REGION Network 105: STATE Num:300 StChkTTPos
   RUNG wire#powerrail
      Contact( #s300_StChkTTPos )
      wire#w1
      I_Contact( #sStWtResetRel )
      I_Contact( #s300_StChkTTPos_T1 )
      I_Contact( #s300_StChkTTPos_T2 )
      I_Contact( #s300_StChkTTPos_T3 )
      wire#w2
      Coil( #s300_StChkTTPos )
   END_RUNG
   RUNG wire#powerrail
      Contact( #s20_StChkForPalletPresent_T4 )
   END_RUNG wire#w1
   RUNG wire#w2
      { S7_GenerateENO := "TRUE" } Move(in := 300, out1 => #StateNo)
   END_RUNG
   // the same network as SCL:
   #s300_StChkTTPos := (#s300_StChkTTPos OR #s20_StChkForPalletPresent_T4) AND NOT #sStWtResetRel AND NOT #s300_StChkTTPos_T1 AND NOT #s300_StChkTTPos_T2 AND NOT #s300_StChkTTPos_T3;
   IF #s300_StChkTTPos THEN #StateNo := 300; END_IF;
END_REGION

REGION Network 106: Actions for STATE Num:300 StChkTTPos
   RUNG wire#powerrail
      Contact( #s300_StChkTTPos )
      Coil( #qOutput1 )
   END_RUNG
   // the same network as SCL:
   #qOutput1 := #s300_StChkTTPos;
END_REGION

REGION Network 107: Transition for STATE Num:310 StWtRTRFrmTTUpAt0
   RUNG wire#powerrail
      Contact( #s310_StWtRTRFrmTTUpAt0 )
      I_Contact( #sStWtResetRel )
      Contact( #sSst )
      wire#w1
      Contact( #sTTUp_Timer_ON.Q )
      Coil( #s310_StWtRTRFrmTTUpAt0_T1 )
   END_RUNG
   RUNG wire#w1
      I_Contact( #s310_StWtRTRFrmTTUpAt0_T1 )
      Contact( #iOTS_Frm_Prev_TTUp )
      I_Contact( #sTTUp_Timer_ON.Q )
      Coil( #s310_StWtRTRFrmTTUpAt0_T2 )
   END_RUNG
   // the same network as SCL:
   #_w1 := #s310_StWtRTRFrmTTUpAt0 AND NOT #sStWtResetRel AND #sSst;
   #s310_StWtRTRFrmTTUpAt0_T1 := #_w1 AND #sTTUp_Timer_ON.Q;
   #s310_StWtRTRFrmTTUpAt0_T2 := #_w1 AND NOT #s310_StWtRTRFrmTTUpAt0_T1 AND #iOTS_Frm_Prev_TTUp AND NOT #sTTUp_Timer_ON.Q;
END_REGION

REGION Network 108: STATE Num:310 StWtRTRFrmTTUpAt0
   RUNG wire#powerrail
      Contact( #s310_StWtRTRFrmTTUpAt0 )
      wire#w1
      I_Contact( #sStWtResetRel )
      I_Contact( #s310_StWtRTRFrmTTUpAt0_T1 )
      I_Contact( #s310_StWtRTRFrmTTUpAt0_T2 )
      wire#w2
      Coil( #s310_StWtRTRFrmTTUpAt0 )
   END_RUNG
   RUNG wire#powerrail
      Contact( #s300_StChkTTPos_T1 )
   END_RUNG wire#w1
   RUNG wire#w2
      { S7_GenerateENO := "TRUE" } Move(in := 310, out1 => #StateNo)
   END_RUNG
   // the same network as SCL:
   #s310_StWtRTRFrmTTUpAt0 := (#s310_StWtRTRFrmTTUpAt0 OR #s300_StChkTTPos_T1) AND NOT #sStWtResetRel AND NOT #s310_StWtRTRFrmTTUpAt0_T1 AND NOT #s310_StWtRTRFrmTTUpAt0_T2;
   IF #s310_StWtRTRFrmTTUpAt0 THEN #StateNo := 310; END_IF;
END_REGION

REGION Network 109: Actions for STATE Num:310 StWtRTRFrmTTUpAt0
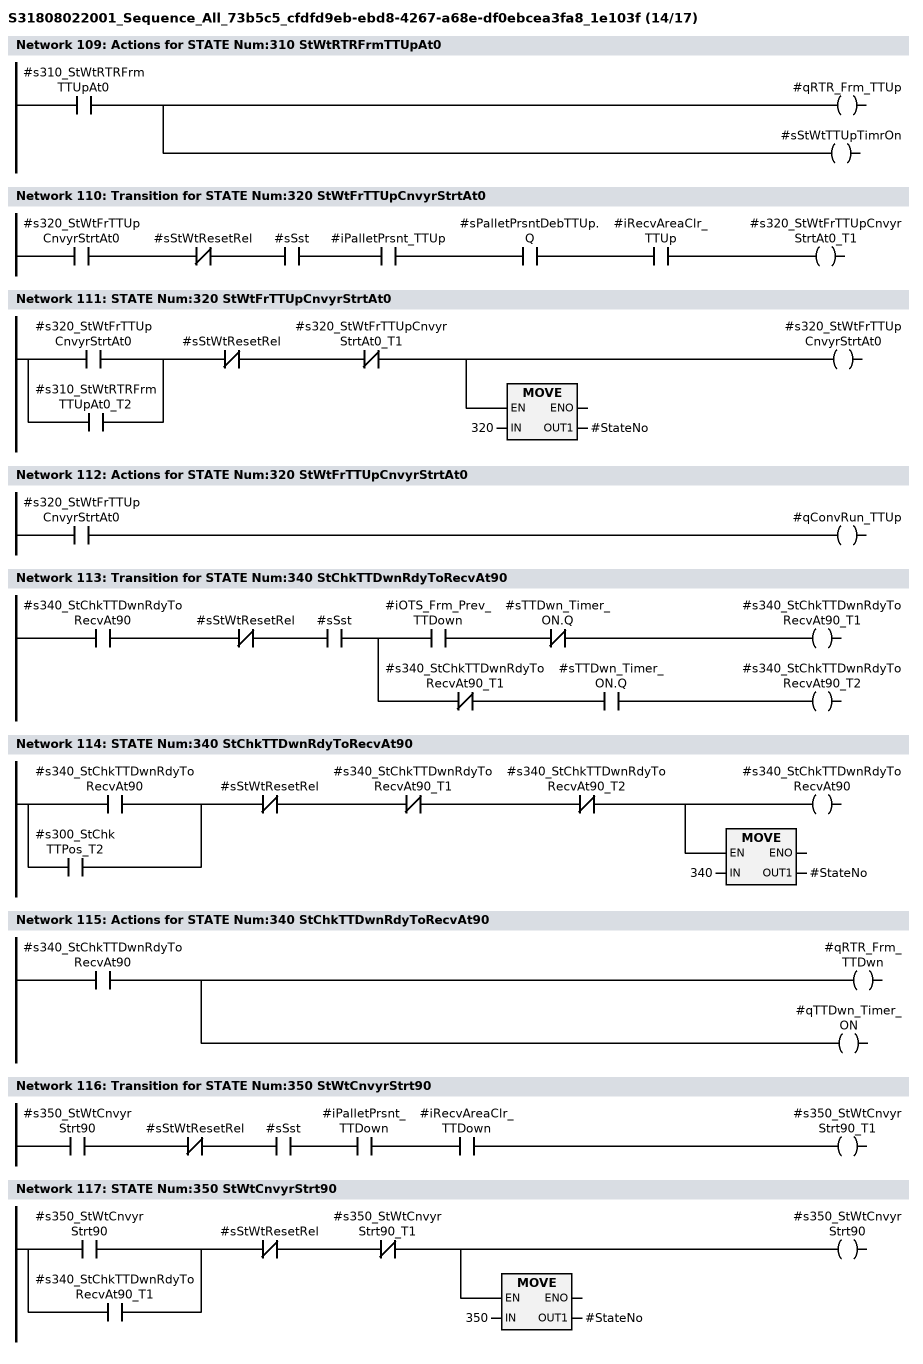
   RUNG wire#powerrail
      Contact( #s310_StWtRTRFrmTTUpAt0 )
      wire#w1
      Coil( #qRTR_Frm_TTUp )
   END_RUNG
   RUNG wire#w1
      Coil( #sStWtTTUpTimrOn )
   END_RUNG
   // the same network as SCL:
   #qRTR_Frm_TTUp := #s310_StWtRTRFrmTTUpAt0;
   #sStWtTTUpTimrOn := #s310_StWtRTRFrmTTUpAt0;
END_REGION

REGION Network 110: Transition for STATE Num:320 StWtFrTTUpCnvyrStrtAt0
   RUNG wire#powerrail
      Contact( #s320_StWtFrTTUpCnvyrStrtAt0 )
      I_Contact( #sStWtResetRel )
      Contact( #sSst )
      Contact( #iPalletPrsnt_TTUp )
      Contact( #sPalletPrsntDebTTUp.Q )
      Contact( #iRecvAreaClr_TTUp )
      Coil( #s320_StWtFrTTUpCnvyrStrtAt0_T1 )
   END_RUNG
   // the same network as SCL:
   #s320_StWtFrTTUpCnvyrStrtAt0_T1 := #s320_StWtFrTTUpCnvyrStrtAt0 AND NOT #sStWtResetRel AND #sSst AND #iPalletPrsnt_TTUp AND #sPalletPrsntDebTTUp.Q AND #iRecvAreaClr_TTUp;
END_REGION

REGION Network 111: STATE Num:320 StWtFrTTUpCnvyrStrtAt0
   RUNG wire#powerrail
      Contact( #s320_StWtFrTTUpCnvyrStrtAt0 )
      wire#w1
      I_Contact( #sStWtResetRel )
      I_Contact( #s320_StWtFrTTUpCnvyrStrtAt0_T1 )
      wire#w2
      Coil( #s320_StWtFrTTUpCnvyrStrtAt0 )
   END_RUNG
   RUNG wire#powerrail
      Contact( #s310_StWtRTRFrmTTUpAt0_T2 )
   END_RUNG wire#w1
   RUNG wire#w2
      { S7_GenerateENO := "TRUE" } Move(in := 320, out1 => #StateNo)
   END_RUNG
   // the same network as SCL:
   #s320_StWtFrTTUpCnvyrStrtAt0 := (#s320_StWtFrTTUpCnvyrStrtAt0 OR #s310_StWtRTRFrmTTUpAt0_T2) AND NOT #sStWtResetRel AND NOT #s320_StWtFrTTUpCnvyrStrtAt0_T1;
   IF #s320_StWtFrTTUpCnvyrStrtAt0 THEN #StateNo := 320; END_IF;
END_REGION

REGION Network 112: Actions for STATE Num:320 StWtFrTTUpCnvyrStrtAt0
   RUNG wire#powerrail
      Contact( #s320_StWtFrTTUpCnvyrStrtAt0 )
      Coil( #qConvRun_TTUp )
   END_RUNG
   // the same network as SCL:
   #qConvRun_TTUp := #s320_StWtFrTTUpCnvyrStrtAt0;
END_REGION

REGION Network 113: Transition for STATE Num:340 StChkTTDwnRdyToRecvAt90
   RUNG wire#powerrail
      Contact( #s340_StChkTTDwnRdyToRecvAt90 )
      I_Contact( #sStWtResetRel )
      Contact( #sSst )
      wire#w1
      Contact( #iOTS_Frm_Prev_TTDown )
      I_Contact( #sTTDwn_Timer_ON.Q )
      Coil( #s340_StChkTTDwnRdyToRecvAt90_T1 )
   END_RUNG
   RUNG wire#w1
      I_Contact( #s340_StChkTTDwnRdyToRecvAt90_T1 )
      Contact( #sTTDwn_Timer_ON.Q )
      Coil( #s340_StChkTTDwnRdyToRecvAt90_T2 )
   END_RUNG
   // the same network as SCL:
   #_w1 := #s340_StChkTTDwnRdyToRecvAt90 AND NOT #sStWtResetRel AND #sSst;
   #s340_StChkTTDwnRdyToRecvAt90_T1 := #_w1 AND #iOTS_Frm_Prev_TTDown AND NOT #sTTDwn_Timer_ON.Q;
   #s340_StChkTTDwnRdyToRecvAt90_T2 := #_w1 AND NOT #s340_StChkTTDwnRdyToRecvAt90_T1 AND #sTTDwn_Timer_ON.Q;
END_REGION

REGION Network 114: STATE Num:340 StChkTTDwnRdyToRecvAt90
   RUNG wire#powerrail
      Contact( #s340_StChkTTDwnRdyToRecvAt90 )
      wire#w1
      I_Contact( #sStWtResetRel )
      I_Contact( #s340_StChkTTDwnRdyToRecvAt90_T1 )
      I_Contact( #s340_StChkTTDwnRdyToRecvAt90_T2 )
      wire#w2
      Coil( #s340_StChkTTDwnRdyToRecvAt90 )
   END_RUNG
   RUNG wire#powerrail
      Contact( #s300_StChkTTPos_T2 )
   END_RUNG wire#w1
   RUNG wire#w2
      { S7_GenerateENO := "TRUE" } Move(in := 340, out1 => #StateNo)
   END_RUNG
   // the same network as SCL:
   #s340_StChkTTDwnRdyToRecvAt90 := (#s340_StChkTTDwnRdyToRecvAt90 OR #s300_StChkTTPos_T2) AND NOT #sStWtResetRel AND NOT #s340_StChkTTDwnRdyToRecvAt90_T1 AND NOT #s340_StChkTTDwnRdyToRecvAt90_T2;
   IF #s340_StChkTTDwnRdyToRecvAt90 THEN #StateNo := 340; END_IF;
END_REGION

REGION Network 115: Actions for STATE Num:340 StChkTTDwnRdyToRecvAt90
   RUNG wire#powerrail
      Contact( #s340_StChkTTDwnRdyToRecvAt90 )
      wire#w1
      Coil( #qRTR_Frm_TTDwn )
   END_RUNG
   RUNG wire#w1
      Coil( #qTTDwn_Timer_ON )
   END_RUNG
   // the same network as SCL:
   #qRTR_Frm_TTDwn := #s340_StChkTTDwnRdyToRecvAt90;
   #qTTDwn_Timer_ON := #s340_StChkTTDwnRdyToRecvAt90;
END_REGION

REGION Network 116: Transition for STATE Num:350 StWtCnvyrStrt90
   RUNG wire#powerrail
      Contact( #s350_StWtCnvyrStrt90 )
      I_Contact( #sStWtResetRel )
      Contact( #sSst )
      Contact( #iPalletPrsnt_TTDown )
      Contact( #iRecvAreaClr_TTDown )
      Coil( #s350_StWtCnvyrStrt90_T1 )
   END_RUNG
   // the same network as SCL:
   #s350_StWtCnvyrStrt90_T1 := #s350_StWtCnvyrStrt90 AND NOT #sStWtResetRel AND #sSst AND #iPalletPrsnt_TTDown AND #iRecvAreaClr_TTDown;
END_REGION

REGION Network 117: STATE Num:350 StWtCnvyrStrt90
   RUNG wire#powerrail
      Contact( #s350_StWtCnvyrStrt90 )
      wire#w1
      I_Contact( #sStWtResetRel )
      I_Contact( #s350_StWtCnvyrStrt90_T1 )
      wire#w2
      Coil( #s350_StWtCnvyrStrt90 )
   END_RUNG
   RUNG wire#powerrail
      Contact( #s340_StChkTTDwnRdyToRecvAt90_T1 )
   END_RUNG wire#w1
   RUNG wire#w2
      { S7_GenerateENO := "TRUE" } Move(in := 350, out1 => #StateNo)
   END_RUNG
   // the same network as SCL:
   #s350_StWtCnvyrStrt90 := (#s350_StWtCnvyrStrt90 OR #s340_StChkTTDwnRdyToRecvAt90_T1) AND NOT #sStWtResetRel AND NOT #s350_StWtCnvyrStrt90_T1;
   IF #s350_StWtCnvyrStrt90 THEN #StateNo := 350; END_IF;
END_REGION

REGION Network 118: Actions for STATE Num:350 StWtCnvyrStrt90
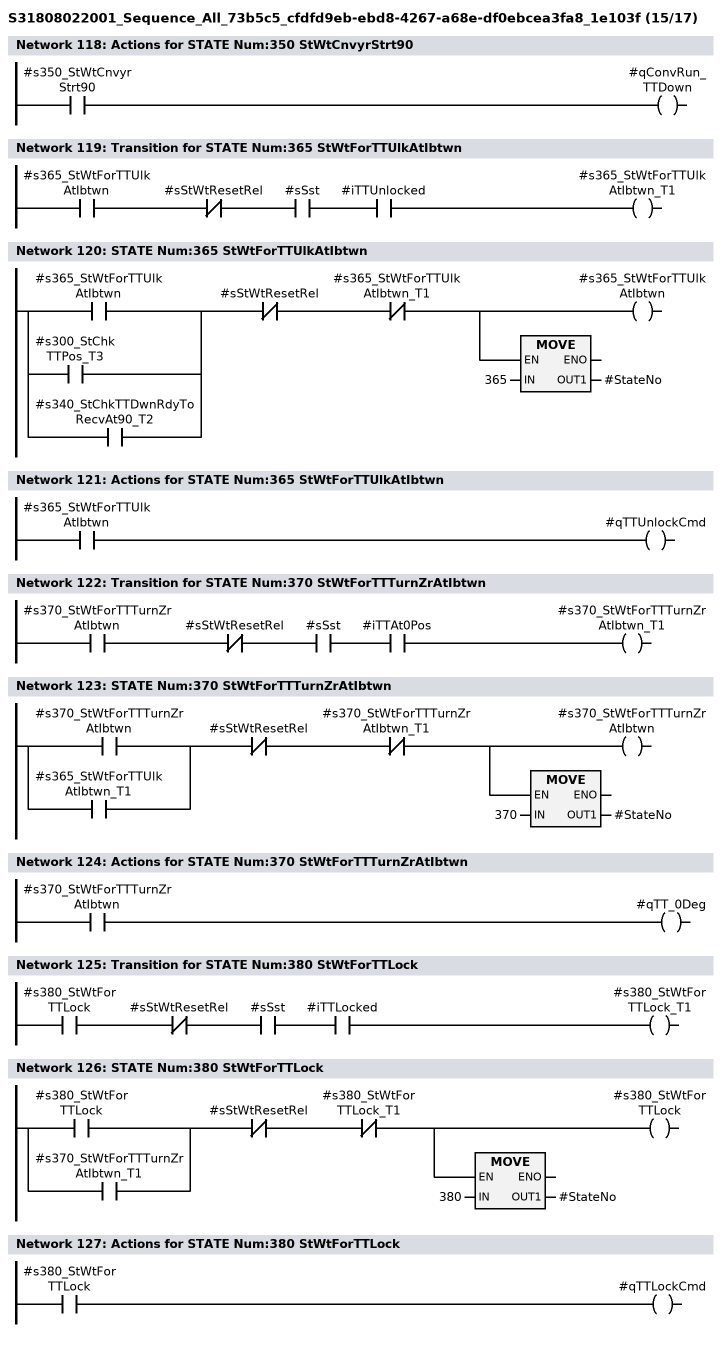
   RUNG wire#powerrail
      Contact( #s350_StWtCnvyrStrt90 )
      Coil( #qConvRun_TTDown )
   END_RUNG
   // the same network as SCL:
   #qConvRun_TTDown := #s350_StWtCnvyrStrt90;
END_REGION

REGION Network 119: Transition for STATE Num:365 StWtForTTUlkAtIbtwn
   RUNG wire#powerrail
      Contact( #s365_StWtForTTUlkAtIbtwn )
      I_Contact( #sStWtResetRel )
      Contact( #sSst )
      Contact( #iTTUnlocked )
      Coil( #s365_StWtForTTUlkAtIbtwn_T1 )
   END_RUNG
   // the same network as SCL:
   #s365_StWtForTTUlkAtIbtwn_T1 := #s365_StWtForTTUlkAtIbtwn AND NOT #sStWtResetRel AND #sSst AND #iTTUnlocked;
END_REGION

REGION Network 120: STATE Num:365 StWtForTTUlkAtIbtwn
   RUNG wire#powerrail
      Contact( #s365_StWtForTTUlkAtIbtwn )
      wire#w1
      I_Contact( #sStWtResetRel )
      I_Contact( #s365_StWtForTTUlkAtIbtwn_T1 )
      wire#w2
      Coil( #s365_StWtForTTUlkAtIbtwn )
   END_RUNG
   RUNG wire#powerrail
      Contact( #s300_StChkTTPos_T3 )
   END_RUNG wire#w1
   RUNG wire#powerrail
      Contact( #s340_StChkTTDwnRdyToRecvAt90_T2 )
   END_RUNG wire#w1
   RUNG wire#w2
      { S7_GenerateENO := "TRUE" } Move(in := 365, out1 => #StateNo)
   END_RUNG
   // the same network as SCL:
   #s365_StWtForTTUlkAtIbtwn := (#s365_StWtForTTUlkAtIbtwn OR #s300_StChkTTPos_T3 OR #s340_StChkTTDwnRdyToRecvAt90_T2) AND NOT #sStWtResetRel AND NOT #s365_StWtForTTUlkAtIbtwn_T1;
   IF #s365_StWtForTTUlkAtIbtwn THEN #StateNo := 365; END_IF;
END_REGION

REGION Network 121: Actions for STATE Num:365 StWtForTTUlkAtIbtwn
   RUNG wire#powerrail
      Contact( #s365_StWtForTTUlkAtIbtwn )
      Coil( #qTTUnlockCmd )
   END_RUNG
   // the same network as SCL:
   #qTTUnlockCmd := #s365_StWtForTTUlkAtIbtwn;
END_REGION

REGION Network 122: Transition for STATE Num:370 StWtForTTTurnZrAtIbtwn
   RUNG wire#powerrail
      Contact( #s370_StWtForTTTurnZrAtIbtwn )
      I_Contact( #sStWtResetRel )
      Contact( #sSst )
      Contact( #iTTAt0Pos )
      Coil( #s370_StWtForTTTurnZrAtIbtwn_T1 )
   END_RUNG
   // the same network as SCL:
   #s370_StWtForTTTurnZrAtIbtwn_T1 := #s370_StWtForTTTurnZrAtIbtwn AND NOT #sStWtResetRel AND #sSst AND #iTTAt0Pos;
END_REGION

REGION Network 123: STATE Num:370 StWtForTTTurnZrAtIbtwn
   RUNG wire#powerrail
      Contact( #s370_StWtForTTTurnZrAtIbtwn )
      wire#w1
      I_Contact( #sStWtResetRel )
      I_Contact( #s370_StWtForTTTurnZrAtIbtwn_T1 )
      wire#w2
      Coil( #s370_StWtForTTTurnZrAtIbtwn )
   END_RUNG
   RUNG wire#powerrail
      Contact( #s365_StWtForTTUlkAtIbtwn_T1 )
   END_RUNG wire#w1
   RUNG wire#w2
      { S7_GenerateENO := "TRUE" } Move(in := 370, out1 => #StateNo)
   END_RUNG
   // the same network as SCL:
   #s370_StWtForTTTurnZrAtIbtwn := (#s370_StWtForTTTurnZrAtIbtwn OR #s365_StWtForTTUlkAtIbtwn_T1) AND NOT #sStWtResetRel AND NOT #s370_StWtForTTTurnZrAtIbtwn_T1;
   IF #s370_StWtForTTTurnZrAtIbtwn THEN #StateNo := 370; END_IF;
END_REGION

REGION Network 124: Actions for STATE Num:370 StWtForTTTurnZrAtIbtwn
   RUNG wire#powerrail
      Contact( #s370_StWtForTTTurnZrAtIbtwn )
      Coil( #qTT_0Deg )
   END_RUNG
   // the same network as SCL:
   #qTT_0Deg := #s370_StWtForTTTurnZrAtIbtwn;
END_REGION

REGION Network 125: Transition for STATE Num:380 StWtForTTLock
   RUNG wire#powerrail
      Contact( #s380_StWtForTTLock )
      I_Contact( #sStWtResetRel )
      Contact( #sSst )
      Contact( #iTTLocked )
      Coil( #s380_StWtForTTLock_T1 )
   END_RUNG
   // the same network as SCL:
   #s380_StWtForTTLock_T1 := #s380_StWtForTTLock AND NOT #sStWtResetRel AND #sSst AND #iTTLocked;
END_REGION

REGION Network 126: STATE Num:380 StWtForTTLock
   RUNG wire#powerrail
      Contact( #s380_StWtForTTLock )
      wire#w1
      I_Contact( #sStWtResetRel )
      I_Contact( #s380_StWtForTTLock_T1 )
      wire#w2
      Coil( #s380_StWtForTTLock )
   END_RUNG
   RUNG wire#powerrail
      Contact( #s370_StWtForTTTurnZrAtIbtwn_T1 )
   END_RUNG wire#w1
   RUNG wire#w2
      { S7_GenerateENO := "TRUE" } Move(in := 380, out1 => #StateNo)
   END_RUNG
   // the same network as SCL:
   #s380_StWtForTTLock := (#s380_StWtForTTLock OR #s370_StWtForTTTurnZrAtIbtwn_T1) AND NOT #sStWtResetRel AND NOT #s380_StWtForTTLock_T1;
   IF #s380_StWtForTTLock THEN #StateNo := 380; END_IF;
END_REGION

REGION Network 127: Actions for STATE Num:380 StWtForTTLock
   RUNG wire#powerrail
      Contact( #s380_StWtForTTLock )
      Coil( #qTTLockCmd )
   END_RUNG
   // the same network as SCL:
   #qTTLockCmd := #s380_StWtForTTLock;
END_REGION

REGION Network 128: Condition1 for STATE Num:400 Wait for all 2 Sub Sequences to complete
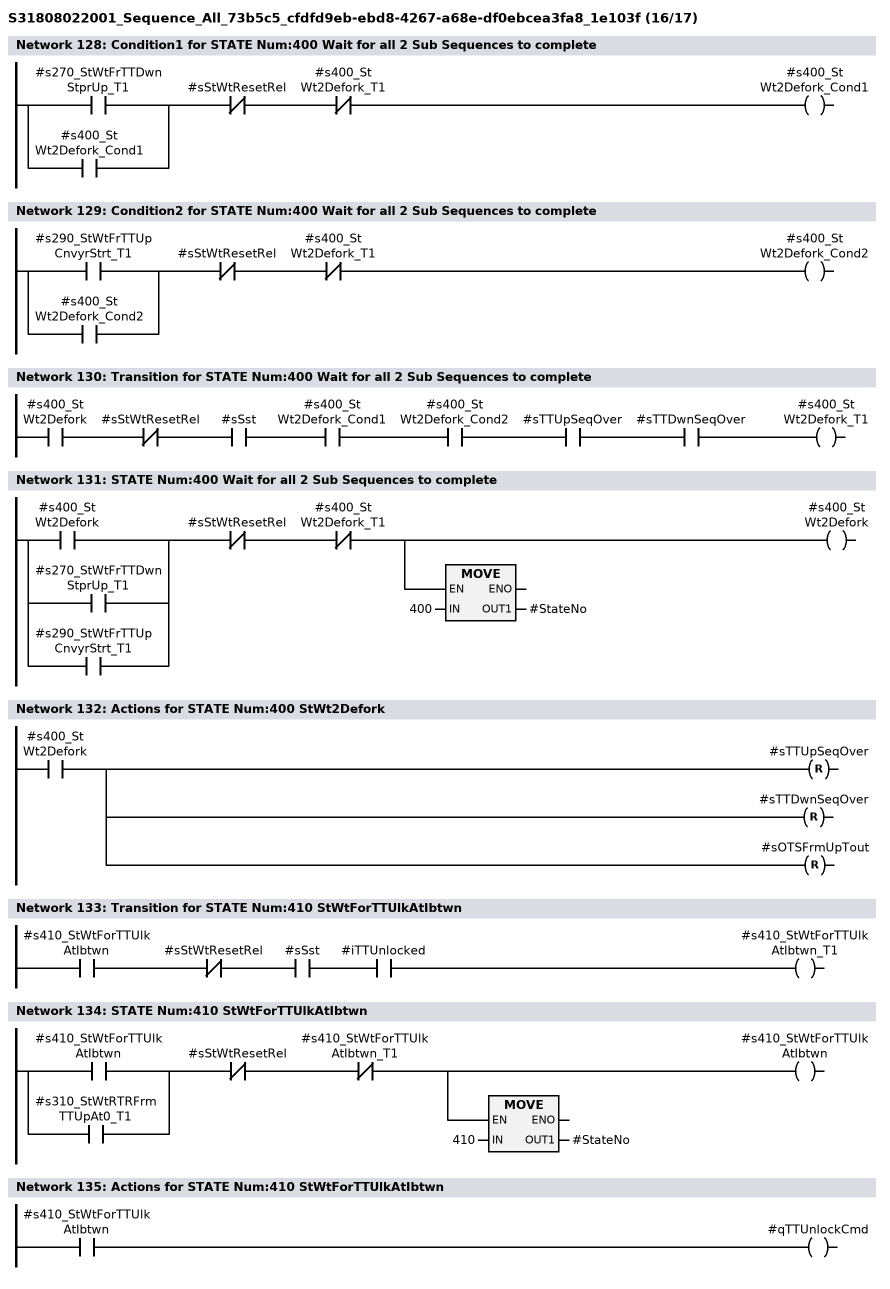
   RUNG wire#powerrail
      Contact( #s270_StWtFrTTDwnStprUp_T1 )
      wire#w1
      I_Contact( #sStWtResetRel )
      I_Contact( #s400_StWt2Defork_T1 )
      Coil( #s400_StWt2Defork_Cond1 )
   END_RUNG
   RUNG wire#powerrail
      Contact( #s400_StWt2Defork_Cond1 )
   END_RUNG wire#w1
   // the same network as SCL:
   #s400_StWt2Defork_Cond1 := (#s270_StWtFrTTDwnStprUp_T1 OR #s400_StWt2Defork_Cond1) AND NOT #sStWtResetRel AND NOT #s400_StWt2Defork_T1;
END_REGION

REGION Network 129: Condition2 for STATE Num:400 Wait for all 2 Sub Sequences to complete
   RUNG wire#powerrail
      Contact( #s290_StWtFrTTUpCnvyrStrt_T1 )
      wire#w1
      I_Contact( #sStWtResetRel )
      I_Contact( #s400_StWt2Defork_T1 )
      Coil( #s400_StWt2Defork_Cond2 )
   END_RUNG
   RUNG wire#powerrail
      Contact( #s400_StWt2Defork_Cond2 )
   END_RUNG wire#w1
   // the same network as SCL:
   #s400_StWt2Defork_Cond2 := (#s290_StWtFrTTUpCnvyrStrt_T1 OR #s400_StWt2Defork_Cond2) AND NOT #sStWtResetRel AND NOT #s400_StWt2Defork_T1;
END_REGION

REGION Network 130: Transition for STATE Num:400 Wait for all 2 Sub Sequences to complete
   RUNG wire#powerrail
      Contact( #s400_StWt2Defork )
      I_Contact( #sStWtResetRel )
      Contact( #sSst )
      Contact( #s400_StWt2Defork_Cond1 )
      Contact( #s400_StWt2Defork_Cond2 )
      Contact( #sTTUpSeqOver )
      Contact( #sTTDwnSeqOver )
      Coil( #s400_StWt2Defork_T1 )
   END_RUNG
   // the same network as SCL:
   #s400_StWt2Defork_T1 := #s400_StWt2Defork AND NOT #sStWtResetRel AND #sSst AND #s400_StWt2Defork_Cond1 AND #s400_StWt2Defork_Cond2 AND #sTTUpSeqOver AND #sTTDwnSeqOver;
END_REGION

REGION Network 131: STATE Num:400 Wait for all 2 Sub Sequences to complete
   RUNG wire#powerrail
      Contact( #s400_StWt2Defork )
      wire#w1
      I_Contact( #sStWtResetRel )
      I_Contact( #s400_StWt2Defork_T1 )
      wire#w2
      Coil( #s400_StWt2Defork )
   END_RUNG
   RUNG wire#powerrail
      Contact( #s270_StWtFrTTDwnStprUp_T1 )
   END_RUNG wire#w1
   RUNG wire#powerrail
      Contact( #s290_StWtFrTTUpCnvyrStrt_T1 )
   END_RUNG wire#w1
   RUNG wire#w2
      { S7_GenerateENO := "TRUE" } Move(in := 400, out1 => #StateNo)
   END_RUNG
   // the same network as SCL:
   #s400_StWt2Defork := (#s400_StWt2Defork OR #s270_StWtFrTTDwnStprUp_T1 OR #s290_StWtFrTTUpCnvyrStrt_T1) AND NOT #sStWtResetRel AND NOT #s400_StWt2Defork_T1;
   IF #s400_StWt2Defork THEN #StateNo := 400; END_IF;
END_REGION

REGION Network 132: Actions for STATE Num:400 StWt2Defork
   RUNG wire#powerrail
      Contact( #s400_StWt2Defork )
      wire#w1
      R_Coil( #sTTUpSeqOver )
   END_RUNG
   RUNG wire#w1
      R_Coil( #sTTDwnSeqOver )
   END_RUNG
   RUNG wire#w1
      R_Coil( #sOTSFrmUpTout )
   END_RUNG
   // the same network as SCL:
   IF #s400_StWt2Defork THEN
       #sTTUpSeqOver := FALSE;
       #sTTDwnSeqOver := FALSE;
       #sOTSFrmUpTout := FALSE;
   END_IF;
END_REGION

REGION Network 133: Transition for STATE Num:410 StWtForTTUlkAtIbtwn
   RUNG wire#powerrail
      Contact( #s410_StWtForTTUlkAtIbtwn )
      I_Contact( #sStWtResetRel )
      Contact( #sSst )
      Contact( #iTTUnlocked )
      Coil( #s410_StWtForTTUlkAtIbtwn_T1 )
   END_RUNG
   // the same network as SCL:
   #s410_StWtForTTUlkAtIbtwn_T1 := #s410_StWtForTTUlkAtIbtwn AND NOT #sStWtResetRel AND #sSst AND #iTTUnlocked;
END_REGION

REGION Network 134: STATE Num:410 StWtForTTUlkAtIbtwn
   RUNG wire#powerrail
      Contact( #s410_StWtForTTUlkAtIbtwn )
      wire#w1
      I_Contact( #sStWtResetRel )
      I_Contact( #s410_StWtForTTUlkAtIbtwn_T1 )
      wire#w2
      Coil( #s410_StWtForTTUlkAtIbtwn )
   END_RUNG
   RUNG wire#powerrail
      Contact( #s310_StWtRTRFrmTTUpAt0_T1 )
   END_RUNG wire#w1
   RUNG wire#w2
      { S7_GenerateENO := "TRUE" } Move(in := 410, out1 => #StateNo)
   END_RUNG
   // the same network as SCL:
   #s410_StWtForTTUlkAtIbtwn := (#s410_StWtForTTUlkAtIbtwn OR #s310_StWtRTRFrmTTUpAt0_T1) AND NOT #sStWtResetRel AND NOT #s410_StWtForTTUlkAtIbtwn_T1;
   IF #s410_StWtForTTUlkAtIbtwn THEN #StateNo := 410; END_IF;
END_REGION

REGION Network 135: Actions for STATE Num:410 StWtForTTUlkAtIbtwn
   RUNG wire#powerrail
      Contact( #s410_StWtForTTUlkAtIbtwn )
      Coil( #qTTUnlockCmd )
   END_RUNG
   // the same network as SCL:
   #qTTUnlockCmd := #s410_StWtForTTUlkAtIbtwn;
END_REGION

REGION Network 136: Transition for STATE Num:415 StWtForTTTurn90AtIbtwn
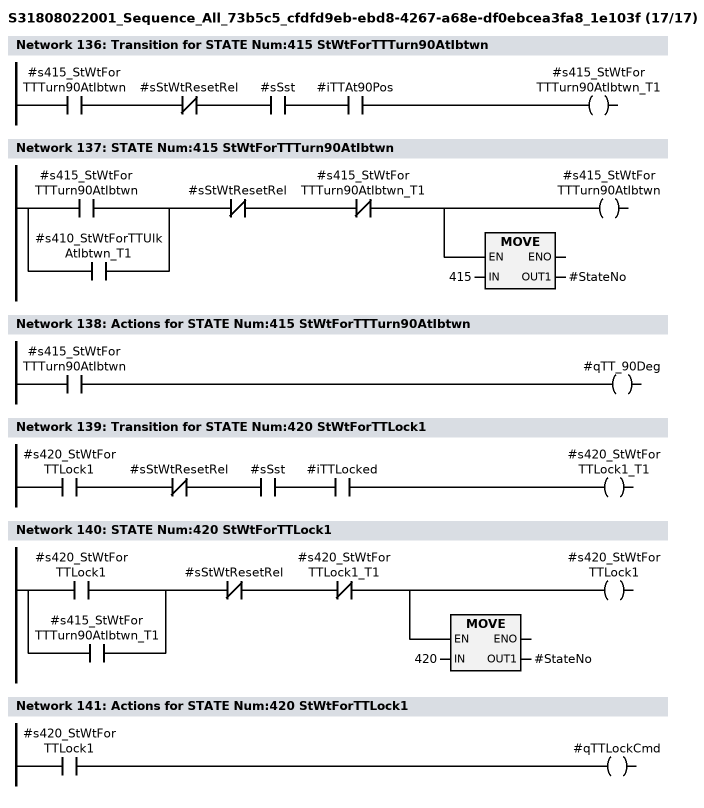
   RUNG wire#powerrail
      Contact( #s415_StWtForTTTurn90AtIbtwn )
      I_Contact( #sStWtResetRel )
      Contact( #sSst )
      Contact( #iTTAt90Pos )
      Coil( #s415_StWtForTTTurn90AtIbtwn_T1 )
   END_RUNG
   // the same network as SCL:
   #s415_StWtForTTTurn90AtIbtwn_T1 := #s415_StWtForTTTurn90AtIbtwn AND NOT #sStWtResetRel AND #sSst AND #iTTAt90Pos;
END_REGION

REGION Network 137: STATE Num:415 StWtForTTTurn90AtIbtwn
   RUNG wire#powerrail
      Contact( #s415_StWtForTTTurn90AtIbtwn )
      wire#w1
      I_Contact( #sStWtResetRel )
      I_Contact( #s415_StWtForTTTurn90AtIbtwn_T1 )
      wire#w2
      Coil( #s415_StWtForTTTurn90AtIbtwn )
   END_RUNG
   RUNG wire#powerrail
      Contact( #s410_StWtForTTUlkAtIbtwn_T1 )
   END_RUNG wire#w1
   RUNG wire#w2
      { S7_GenerateENO := "TRUE" } Move(in := 415, out1 => #StateNo)
   END_RUNG
   // the same network as SCL:
   #s415_StWtForTTTurn90AtIbtwn := (#s415_StWtForTTTurn90AtIbtwn OR #s410_StWtForTTUlkAtIbtwn_T1) AND NOT #sStWtResetRel AND NOT #s415_StWtForTTTurn90AtIbtwn_T1;
   IF #s415_StWtForTTTurn90AtIbtwn THEN #StateNo := 415; END_IF;
END_REGION

REGION Network 138: Actions for STATE Num:415 StWtForTTTurn90AtIbtwn
   RUNG wire#powerrail
      Contact( #s415_StWtForTTTurn90AtIbtwn )
      Coil( #qTT_90Deg )
   END_RUNG
   // the same network as SCL:
   #qTT_90Deg := #s415_StWtForTTTurn90AtIbtwn;
END_REGION

REGION Network 139: Transition for STATE Num:420 StWtForTTLock1
   RUNG wire#powerrail
      Contact( #s420_StWtForTTLock1 )
      I_Contact( #sStWtResetRel )
      Contact( #sSst )
      Contact( #iTTLocked )
      Coil( #s420_StWtForTTLock1_T1 )
   END_RUNG
   // the same network as SCL:
   #s420_StWtForTTLock1_T1 := #s420_StWtForTTLock1 AND NOT #sStWtResetRel AND #sSst AND #iTTLocked;
END_REGION

REGION Network 140: STATE Num:420 StWtForTTLock1
   RUNG wire#powerrail
      Contact( #s420_StWtForTTLock1 )
      wire#w1
      I_Contact( #sStWtResetRel )
      I_Contact( #s420_StWtForTTLock1_T1 )
      wire#w2
      Coil( #s420_StWtForTTLock1 )
   END_RUNG
   RUNG wire#powerrail
      Contact( #s415_StWtForTTTurn90AtIbtwn_T1 )
   END_RUNG wire#w1
   RUNG wire#w2
      { S7_GenerateENO := "TRUE" } Move(in := 420, out1 => #StateNo)
   END_RUNG
   // the same network as SCL:
   #s420_StWtForTTLock1 := (#s420_StWtForTTLock1 OR #s415_StWtForTTTurn90AtIbtwn_T1) AND NOT #sStWtResetRel AND NOT #s420_StWtForTTLock1_T1;
   IF #s420_StWtForTTLock1 THEN #StateNo := 420; END_IF;
END_REGION

REGION Network 141: Actions for STATE Num:420 StWtForTTLock1
   RUNG wire#powerrail
      Contact( #s420_StWtForTTLock1 )
      Coil( #qTTLockCmd )
   END_RUNG
   // the same network as SCL:
   #qTTLockCmd := #s420_StWtForTTLock1;
END_REGION
END_FUNCTION_BLOCK

ORGANIZATION_BLOCK "Main"   // OB1, LAD, ProgramCycle
TITLE = "Main Program Sweep (Cycle)"
{ S7_Optimized_Access := 'TRUE' }
VERSION : 0.1
   VAR_INPUT
      Initial_Call : Bool;   // Initial call of this OB
      Remanence : Bool;   // =True, if remanent data are available
   END_VAR
   VAR_TEMP
      OB1_EV_CLASS : Byte;   // Bits 0-3 = 1 (Coming event), Bits 4-7 = 1 (Event class 1)
      OB1_SCAN_1 : Byte;   // 1 (Cold restart scan 1 of OB 1), 3 (Scan 2-n of OB 1)
      OB1_PRIORITY : Byte;   // Priority of OB Execution
      OB1_OB_NUMBR : Byte;   // 1 (Organization block 1, OB1)
      OB1_RESERVED_1 : Byte;   // Reserved for system
      OB1_RESERVED_2 : Byte;   // Reserved for system
      OB1_PREV_CYCLE : Int;   // Cycle time of previous OB1 scan (milliseconds)
      OB1_MIN_CYCLE : Int;   // Minimum cycle time of OB1 (milliseconds)
      OB1_MAX_CYCLE : Int;   // Maximum cycle time of OB1 (milliseconds)
      OB1_DATE_TIME : Date_And_Time;   // Date and time OB1 started
   END_VAR
BEGIN
END_ORGANIZATION_BLOCK